(* Simple Raw ADC Sensor Reading to Temperature Conversion *)

PROGRAM main
  VAR
    RawADC : REAL;
    Temp : REAL;
    DivInter : REAL;
    MulInter : REAL;
  END_VAR
  VAR  (* added by the conversion: wires and edge detectors of the diagram *)
    _SUB5_OUT : REAL;
  END_VAR

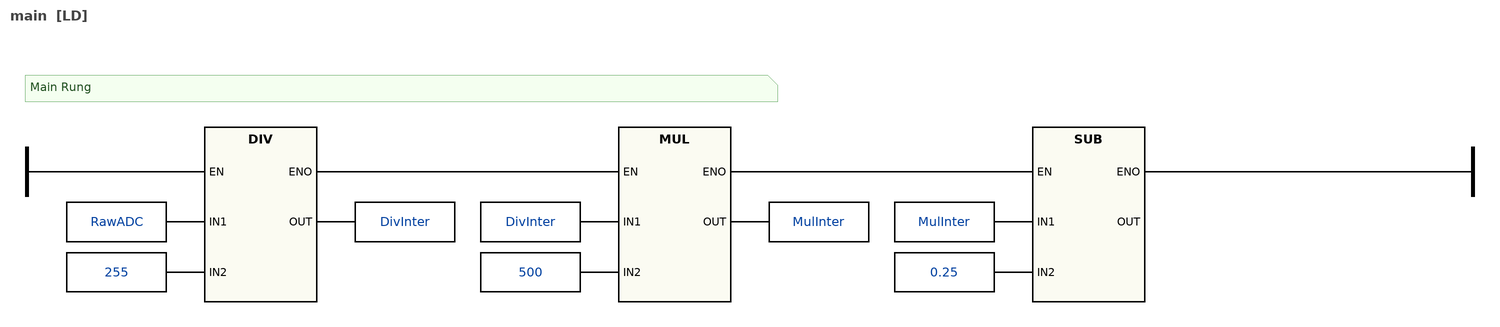
(* LD diagram, written out as Structured Text *)
(* Main Rung *)
DivInter := RawADC / 255;
MulInter := DivInter * 500;
_SUB5_OUT := MulInter - 0.25;
END_PROGRAM
